(* IEC 61131-3 sources: IEC61131-3_ST_SCL_Mutation_Generator/Tests/mutatedCode_timer, 4 files *)

(* ---- M182.st ---- *)
FUNCTION_BLOCK TON_Example

VAR
    StartButton : BOOL;
    Motor       : BOOL;
    StartTimer  : TON;
END_VAR

StartTimer(
    IN := Motor,
 (* MUTATED: VAR_REPLACE *)
    PT := T#5s
);

Motor := StartTimer.Q;

END_FUNCTION_BLOCK

(* ---- M183.st ---- *)
FUNCTION_BLOCK TON_Example

VAR
    StartButton : BOOL;
    Motor       : BOOL;
    StartTimer  : TON;
END_VAR

StartTimer(
    IN := StartButton,
    PT := T#5s
);

StartButton := StartTimer.Q;
 (* MUTATED: VAR_REPLACE *)

END_FUNCTION_BLOCK

(* ---- M184.st ---- *)
FUNCTION_BLOCK TON_Example

VAR
    StartButton : BOOL;
    Motor       : BOOL;
    StartTimer  : TON;
END_VAR

StartTimer(
    IN := StartButton,
    PT := T#5s
);

Motor := NOT (StartTimer.Q);
 (* MUTATED: ASSIGN_NEGATE *)

END_FUNCTION_BLOCK

(* ---- M185.st ---- *)
FUNCTION_BLOCK TON_Example

VAR
    StartButton : BOOL;
    Motor       : BOOL;
    StartTimer  : TON;
END_VAR

StartTimer(
    IN := StartButton,
    PT := T#5s
);

Motor := StartButton; (* MUTATION: TIMER_BYPASS on StartTimer *)

END_FUNCTION_BLOCK
